// SIMATIC STEP 7 (V5.x) project exercice12
// CPU: CPU 314
// station: Matériel
// station: SIMATIC 300(1)
// station: P_ADR_BUS
// program: Programme S7(1)

SYMBOL_TABLE
"START"	I 0.0	BOOL
"ROUGE"	Q 0.0	BOOL
"ORANGE"	Q 0.1	BOOL
"VERT"	Q 0.2	BOOL
END_SYMBOL_TABLE

ORGANIZATION_BLOCK OB 1
TITLE = "Main Program Sweep (Cycle)"
VERSION : 0.1
VAR_TEMP
  OB1_EV_CLASS : BYTE ;	//Bits 0-3 = 1 (Coming event), Bits 4-7 = 1 (Event class 1)
  OB1_SCAN_1 : BYTE ;	//1 (Cold restart scan 1 of OB 1), 3 (Scan 2-n of OB 1)
  OB1_PRIORITY : BYTE ;	//Priority of OB Execution
  OB1_OB_NUMBR : BYTE ;	//1 (Organization block 1, OB1)
  OB1_RESERVED_1 : BYTE ;	//Reserved for system
  OB1_RESERVED_2 : BYTE ;	//Reserved for system
  OB1_PREV_CYCLE : INT ;	//Cycle time of previous OB1 scan (milliseconds)
  OB1_MIN_CYCLE : INT ;	//Minimum cycle time of OB1 (milliseconds)
  OB1_MAX_CYCLE : INT ;	//Maximum cycle time of OB1 (milliseconds)
  OB1_DATE_TIME : DATE_AND_TIME ;	//Date and time OB1 started
END_VAR
BEGIN
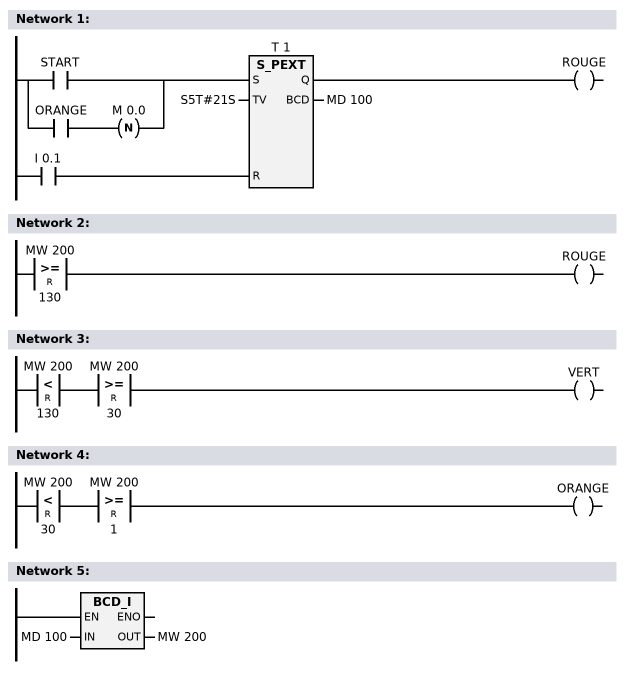
NETWORK
TITLE =
      A(;
      O     "START";
      O(;
      A     "ORANGE";
      BLD   100;
      FN    M 0.0;
      );
      );
      L     S5T#21S;
      SE    T 1;
      A     I 0.1;
      R     T 1;
      NOP   0;
      LC    T 1;
      T     MD 100;
      A     T 1;
      =     "ROUGE";
NETWORK
TITLE =
      L     MW 200;
      L     130;
      >=R;
      =     "ROUGE";
NETWORK
TITLE =
      A(;
      L     MW 200;
      L     130;
      <R;
      );
      A(;
      L     MW 200;
      L     30;
      >=R;
      );
      =     "VERT";
NETWORK
TITLE =
      A(;
      L     MW 200;
      L     30;
      <R;
      );
      A(;
      L     MW 200;
      L     1;
      >=R;
      );
      =     "ORANGE";
NETWORK
TITLE =
      L     MD 100;
      BTI;
      T     MW 200;
      NOP   0;
END_ORGANIZATION_BLOCK
